(* IEC 61131-3 sources: model-first-plc-agent-ai/results/T4-W-04, 2 files *)

(* ---- a1_code.st ---- *)
FUNCTION_BLOCK LevelControlRuntime
VAR_INPUT
    StartCommand : BOOL;
    StopCommand : BOOL;
    LevelMeter : INT;
    FullScaleValue : INT;
    h_span : REAL;
    h_sp : REAL;
    h_target : REAL;
    h_max : REAL;
    eps : REAL;
    t_h : TIME;
    Kp : REAL;
    Ti : REAL;
    Td : REAL;
    CycleTime : TIME;
END_VAR
VAR_OUTPUT
    fill_valve : BOOL;
    discharge_valve : BOOL;
    pid_percent : REAL;
END_VAR
VAR
    StartEdge : R_TRIG;
    SettlingTimer : TON;

    start : BOOL;
    stop : BOOL;
    settled : BOOL;

    (* Region encoding: 0 = LOW, 1 = MID, 2 = HIGH. *)
    r : INT;

    x0 : BOOL := TRUE;
    x1 : BOOL := FALSE;
    WasActive : BOOL := FALSE;

    h : REAL;
    e : REAL;
    CycleSeconds : REAL;

    IntegralTerm : REAL := 0.0;
    IntegralCandidate : REAL;
    PreviousError : REAL := 0.0;
    ProportionalTerm : REAL;
    DerivativeTerm : REAL;
    UnboundedDemand : REAL;
END_VAR

StartEdge(CLK := StartCommand);
start := StartEdge.Q;
stop := StopCommand;

h := INT_TO_REAL(LevelMeter) * h_span / INT_TO_REAL(FullScaleValue);
e := h_sp - h;

IF h < h_target THEN
    r := 0;
ELSIF h < h_max THEN
    r := 1;
ELSE
    r := 2;
END_IF;

CycleSeconds := TIME_TO_REAL(CycleTime) / 1000.0;

(* The non-retentive timer measures continuous time in tolerance
   while x1 is active, not merely the age of x1. *)
SettlingTimer(
    IN := x1 AND (ABS(e) <= eps),
    PT := t_h
);
settled := SettlingTimer.Q;

WasActive := x1;

(* Evaluate transitions from the situation at the start of this scan.
   At most one transition is fired per scan. *)
IF x0 THEN
    IF start AND NOT stop AND NOT (r = 2) THEN
        x0 := FALSE;
        x1 := TRUE;
    END_IF;
ELSIF x1 THEN
    IF stop OR settled OR (r = 2) THEN
        x1 := FALSE;
        x0 := TRUE;
    END_IF;
END_IF;

fill_valve := x1;
discharge_valve := x1;

IF x1 THEN
    (* Initialize controller history on entry to regulation. *)
    IF NOT WasActive THEN
        IntegralTerm := 0.0;
        PreviousError := e;
    END_IF;

    ProportionalTerm := Kp * e;
    DerivativeTerm := 0.0;

    IF (CycleSeconds > 0.0) AND (Td > 0.0) THEN
        DerivativeTerm :=
            Kp * Td * (e - PreviousError) / CycleSeconds;
    END_IF;

    (* Positional PID, with output expressed in percent.
       First test the demand using the existing integral state. *)
    UnboundedDemand :=
        ProportionalTerm + IntegralTerm + DerivativeTerm;

    IF (UnboundedDemand >= 0.0)
        AND (UnboundedDemand <= 100.0)
        AND (Ti > 0.0)
        AND (CycleSeconds > 0.0) THEN

        IntegralCandidate :=
            IntegralTerm + Kp * e * CycleSeconds / Ti;

        UnboundedDemand :=
            ProportionalTerm + IntegralCandidate + DerivativeTerm;

        (* Commit integration only if the resulting output is not
           clamped. Otherwise retain the previous integral state. *)
        IF (UnboundedDemand >= 0.0)
            AND (UnboundedDemand <= 100.0) THEN
            IntegralTerm := IntegralCandidate;
        END_IF;
    END_IF;

    IF UnboundedDemand < 0.0 THEN
        pid_percent := 0.0;
    ELSIF UnboundedDemand > 100.0 THEN
        pid_percent := 100.0;
    ELSE
        pid_percent := UnboundedDemand;
    END_IF;

    PreviousError := e;
ELSE
    pid_percent := 0.0;
    IntegralTerm := 0.0;
    PreviousError := e;

    (* Clear the owned condition immediately on leaving x1. *)
    SettlingTimer(IN := FALSE, PT := t_h);
    settled := FALSE;
END_IF;

END_FUNCTION_BLOCK

PROGRAM Main
VAR
    StartCommand AT %IX100.0 : BOOL;
    StopCommand AT %IX100.1 : BOOL;
    LevelMeter AT %IW100 : INT;
    FillValve AT %QW100 : INT;
    DischargeValve AT %QW101 : INT;
END_VAR
VAR CONSTANT
    FULL_SCALE : INT := 1000;
END_VAR
VAR
    Controller : LevelControlRuntime;

    h_span : REAL := 10.0;
    h_sp : REAL;
    h_target : REAL;
    h_max : REAL;
    eps : REAL;
    t_h : TIME := T#10s;

    (* Initial tuning values; commission for the actual plant.
       Kp units: percent per level unit; Ti and Td units: seconds. *)
    Kp : REAL := 10.0;
    Ti : REAL := 10.0;
    Td : REAL := 0.0;

    CycleTime : TIME := T#20ms;
END_VAR

h_sp := 0.8 * h_span;
h_target := h_sp;
h_max := 0.9 * h_span;
eps := 0.02 * h_span;

Controller(
    StartCommand := StartCommand,
    StopCommand := StopCommand,
    LevelMeter := LevelMeter,
    FullScaleValue := FULL_SCALE,
    h_span := h_span,
    h_sp := h_sp,
    h_target := h_target,
    h_max := h_max,
    eps := eps,
    t_h := t_h,
    Kp := Kp,
    Ti := Ti,
    Td := Td,
    CycleTime := CycleTime
);

IF Controller.fill_valve THEN
    FillValve := REAL_TO_INT(
        Controller.pid_percent * INT_TO_REAL(FULL_SCALE) / 100.0
    );
ELSE
    FillValve := 0;
END_IF;

IF Controller.discharge_valve THEN
    DischargeValve := REAL_TO_INT(0.4 * INT_TO_REAL(FULL_SCALE));
ELSE
    DischargeValve := 0;
END_IF;

END_PROGRAM

CONFIGURATION Config
    RESOURCE PLCResource ON PLC
        TASK ControlTask(INTERVAL := T#20ms, PRIORITY := 0);
        PROGRAM MainInstance WITH ControlTask : Main;
    END_RESOURCE
END_CONFIGURATION

(* ---- a2_code.st ---- *)
FUNCTION_BLOCK FB_LevelControl
VAR_INPUT
    StartCommand : BOOL;
    StopCommand : BOOL;
    LevelMeter : INT;
    h_span : REAL := 10.0;
    Kp : REAL := 10.0;
    Ti : REAL := 10.0;
    Td : REAL := 0.0;
    t_h : TIME := T#10s;
    cycle_seconds : REAL := 0.02;
END_VAR
VAR_OUTPUT
    FillValve : INT;
    DischargeValve : INT;
    fill_valve : BOOL;
    discharge_valve : BOOL;
END_VAR
VAR CONSTANT
    FULL_SCALE : INT := 1000;
    REGION_LOW : INT := 0;
    REGION_MIDDLE : INT := 1;
    REGION_HIGH : INT := 2;
END_VAR
VAR
    StartEdge : R_TRIG;
    HoldTimer : TON;
    start : BOOL;
    stop : BOOL;
    settled : BOOL;
    r : INT;
    sequence_state : INT := 0;
    x0 : BOOL := TRUE;
    x1 : BOOL := FALSE;
    h : REAL;
    h_sp : REAL;
    h_target : REAL;
    h_max : REAL;
    eps : REAL;
    e : REAL;
    previous_error : REAL := 0.0;
    derivative_ready : BOOL := FALSE;
    proportional_term : REAL;
    integral_term : REAL := 0.0;
    derivative_term : REAL;
    integral_candidate : REAL;
    demand_candidate : REAL;
    raw_demand : REAL;
    bounded_demand : REAL;
END_VAR

StartEdge(CLK := StartCommand);
start := StartEdge.Q;
stop := StopCommand;

h := INT_TO_REAL(LevelMeter) * h_span / INT_TO_REAL(FULL_SCALE);
h_sp := 0.8 * h_span;
h_target := h_sp;
h_max := 0.9 * h_span;
eps := 0.02 * h_span;
e := h_sp - h;

IF h < h_target THEN
    r := REGION_LOW;
ELSIF h < h_max THEN
    r := REGION_MIDDLE;
ELSE
    r := REGION_HIGH;
END_IF;

HoldTimer(
    IN := (sequence_state = 1) AND NOT stop
          AND (r <> REGION_HIGH) AND (ABS(e) <= eps),
    PT := t_h
);
settled := HoldTimer.Q;

IF stop THEN
    sequence_state := 0;
ELSE
    CASE sequence_state OF
        0:
            IF start AND (r <> REGION_HIGH) THEN
                sequence_state := 1;
            END_IF;
        1:
            IF settled OR (r = REGION_HIGH) THEN
                sequence_state := 0;
            END_IF;
    ELSE
        sequence_state := 0;
    END_CASE;
END_IF;

x0 := sequence_state = 0;
x1 := sequence_state = 1;
fill_valve := x1;
discharge_valve := x1;

FillValve := 0;
DischargeValve := 0;

IF x1 THEN
    proportional_term := Kp * e;
    derivative_term := 0.0;

    IF derivative_ready AND (cycle_seconds > 0.0) THEN
        derivative_term :=
            Kp * Td * (e - previous_error) / cycle_seconds;
    END_IF;

    raw_demand := proportional_term + integral_term + derivative_term;

    (* Suspend integration whenever the PID demand is clamped.
       Reject an integral increment that would itself cause clamping. *)
    IF (raw_demand >= 0.0) AND (raw_demand <= 100.0)
       AND (Ti > 0.0) AND (cycle_seconds > 0.0) THEN
        integral_candidate :=
            integral_term + Kp * e * cycle_seconds / Ti;
        demand_candidate :=
            proportional_term + integral_candidate + derivative_term;

        IF (demand_candidate >= 0.0)
           AND (demand_candidate <= 100.0) THEN
            integral_term := integral_candidate;
            raw_demand := demand_candidate;
        END_IF;
    END_IF;

    IF raw_demand < 0.0 THEN
        bounded_demand := 0.0;
    ELSIF raw_demand > 100.0 THEN
        bounded_demand := 100.0;
    ELSE
        bounded_demand := raw_demand;
    END_IF;

    FillValve := REAL_TO_INT(
        bounded_demand * INT_TO_REAL(FULL_SCALE) / 100.0
    );
    DischargeValve := REAL_TO_INT(0.4 * INT_TO_REAL(FULL_SCALE));

    previous_error := e;
    derivative_ready := TRUE;
ELSE
    integral_term := 0.0;
    previous_error := e;
    derivative_ready := FALSE;
    bounded_demand := 0.0;
END_IF;

END_FUNCTION_BLOCK

PROGRAM Main
VAR
    StartCommand AT %IX100.0 : BOOL;
    StopCommand AT %IX100.1 : BOOL;
    LevelMeter AT %IW100 : INT;
    FillValve AT %QW100 : INT;
    DischargeValve AT %QW101 : INT;
END_VAR
VAR
    LevelController : FB_LevelControl;
    h_span : REAL := 10.0;
    Kp : REAL := 10.0;
    Ti : REAL := 10.0;
    Td : REAL := 0.0;
    t_h : TIME := T#10s;
END_VAR

(* Kp uses percent opening per level unit; Ti and Td use seconds.
   Initial gain values are commissioning defaults, not tuned plant gains. *)
LevelController(
    StartCommand := StartCommand,
    StopCommand := StopCommand,
    LevelMeter := LevelMeter,
    h_span := h_span,
    Kp := Kp,
    Ti := Ti,
    Td := Td,
    t_h := t_h,
    cycle_seconds := 0.02
);

FillValve := LevelController.FillValve;
DischargeValve := LevelController.DischargeValve;

END_PROGRAM

CONFIGURATION Config0
    RESOURCE Res0 ON PLC
        TASK ControlTask(INTERVAL := T#20ms, PRIORITY := 0);
        PROGRAM MainInstance WITH ControlTask : Main;
    END_RESOURCE
END_CONFIGURATION
